(* IEC 61131-3 sources: codesys-framework/txt/application/WeVe Utils (library)/TimeStamp/I_TimeStampService/Commands, 5 files *)

(* ---- ForceNTPTimeSync.method.st ---- *)
METHOD ForceNTPTimeSync : E_TaskStatus
VAR_INPUT
END_VAR

(* ---- SetLocalTime.method.st ---- *)
METHOD SetLocalTime : E_TaskStatus
VAR_INPUT
	uiYear 					: UINT;
	uiMonth 				: UINT;
	uiDay 					: UINT;
	uiHour 					: UINT;
	uiMinute 				: UINT;
	uiSecond 				: UINT;
END_VAR

(* ---- SetLocalTimeZone.method.st ---- *)
METHOD SetLocalTimeZone : E_TaskStatus
VAR_INPUT
	eTimeZone	: E_TimeZone;
END_VAR

(* ---- SetTimeBase.method.st ---- *)
METHOD SetTimeBase : E_TaskStatus
VAR_INPUT
	eTimeBase : E_TimeBase;
END_VAR

(* ---- SetTimeServer.method.st ---- *)
METHOD SetTimeServer : E_TaskStatus
VAR_INPUT
END_VAR
